// SIMATIC S7-200 project (STEP 7-Micro/WIN), CPU 224XP CN REL 02.01

SYMBOL_TABLE USUARIO1
C_1              VD100
C_0              VD110
L_k              VD180
r_k              VD190
m_k              VD120
m_k_1            VD130
m_k_2            VD140
e_k              VD300
e_k_1            VD160
e_k_2            VD170
Aa               VD200
Bb               VD210
Cc               VD220
Dd               VD230
Ee               VD240
r_k_1            VD250
END_SYMBOL_TABLE

ORGANIZATION_BLOCK PRINCIPAL:OB1
TITLE=COMENTARIOS DEL PROGRAMA
BEGIN
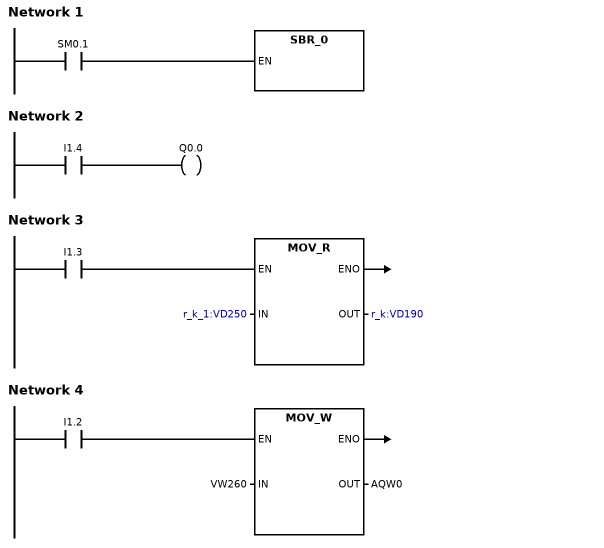
Network 1
LD     SM0.1
CALL   SBR_0:SBR0
Network 2
LD     I1.4
=      Q0.0
Network 3
LD     I1.3
MOVR   r_k_1:VD250, r_k:VD190
Network 4
LD     I1.2
MOVW   VW260, AQW0
END_ORGANIZATION_BLOCK

SUBROUTINE_BLOCK SBR_0:SBR0
TITLE=COMENTARIOS DE LA SUBRUTINA
BEGIN
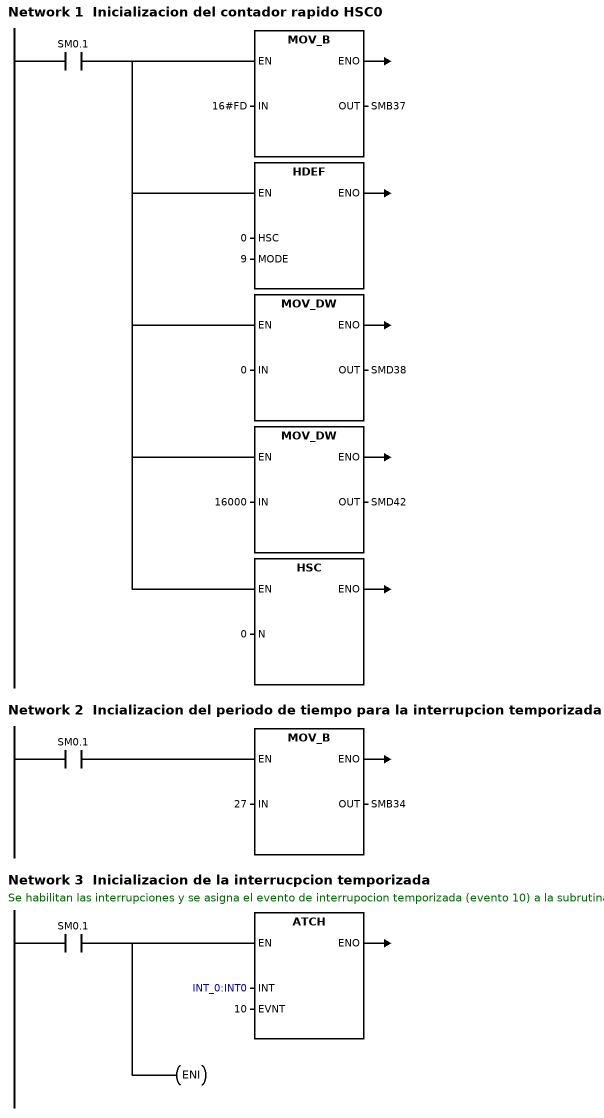
Network 1 // Inicializacion del contador rapido HSC0
LD     SM0.1
MOVB   16#FD, SMB37
HDEF   0, 9
MOVD   0, SMD38
MOVD   16000, SMD42
HSC    0
Network 2 // Incializacion del periodo de tiempo para la interrupcion temporizada
LD     SM0.1
MOVB   27, SMB34
Network 3 // Inicializacion de la interrucpcion temporizada
// Se habilitan las interrupciones y se asigna el evento de interrupocion temporizada (evento 10) a la subrutina de interrupcion INT_0
LD     SM0.1
ATCH   INT_0:INT0, 10
ENI
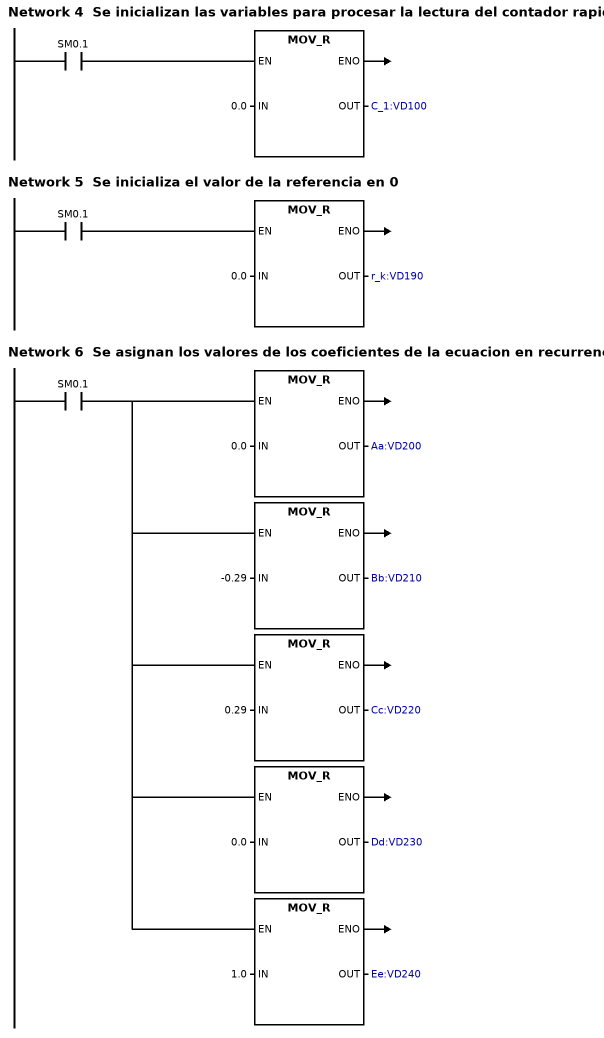
Network 4 // Se inicializan las variables para procesar la lectura del contador rapido HSC0
LD     SM0.1
MOVR   0.0, C_1:VD100
Network 5 // Se inicializa el valor de la referencia en 0
LD     SM0.1
MOVR   0.0, r_k:VD190
Network 6 // Se asignan los valores de los coeficientes de la ecuacion en recurrencia
LD     SM0.1
MOVR   0.0, Aa:VD200
MOVR   -0.29, Bb:VD210
MOVR   0.29, Cc:VD220
MOVR   0.0, Dd:VD230
MOVR   1.0, Ee:VD240
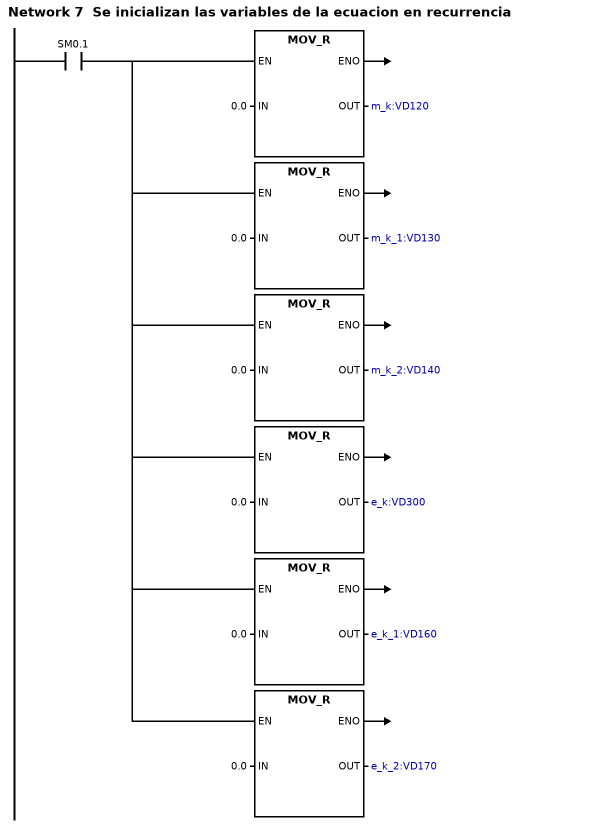
Network 7 // Se inicializan las variables de la ecuacion en recurrencia
LD     SM0.1
MOVR   0.0, m_k:VD120
MOVR   0.0, m_k_1:VD130
MOVR   0.0, m_k_2:VD140
MOVR   0.0, e_k:VD300
MOVR   0.0, e_k_1:VD160
MOVR   0.0, e_k_2:VD170
END_SUBROUTINE_BLOCK

INTERRUPT_BLOCK INT_0:INT0
TITLE=COMENTARIOS DE LA RUTINA DE INTERRUPCIÓN
BEGIN
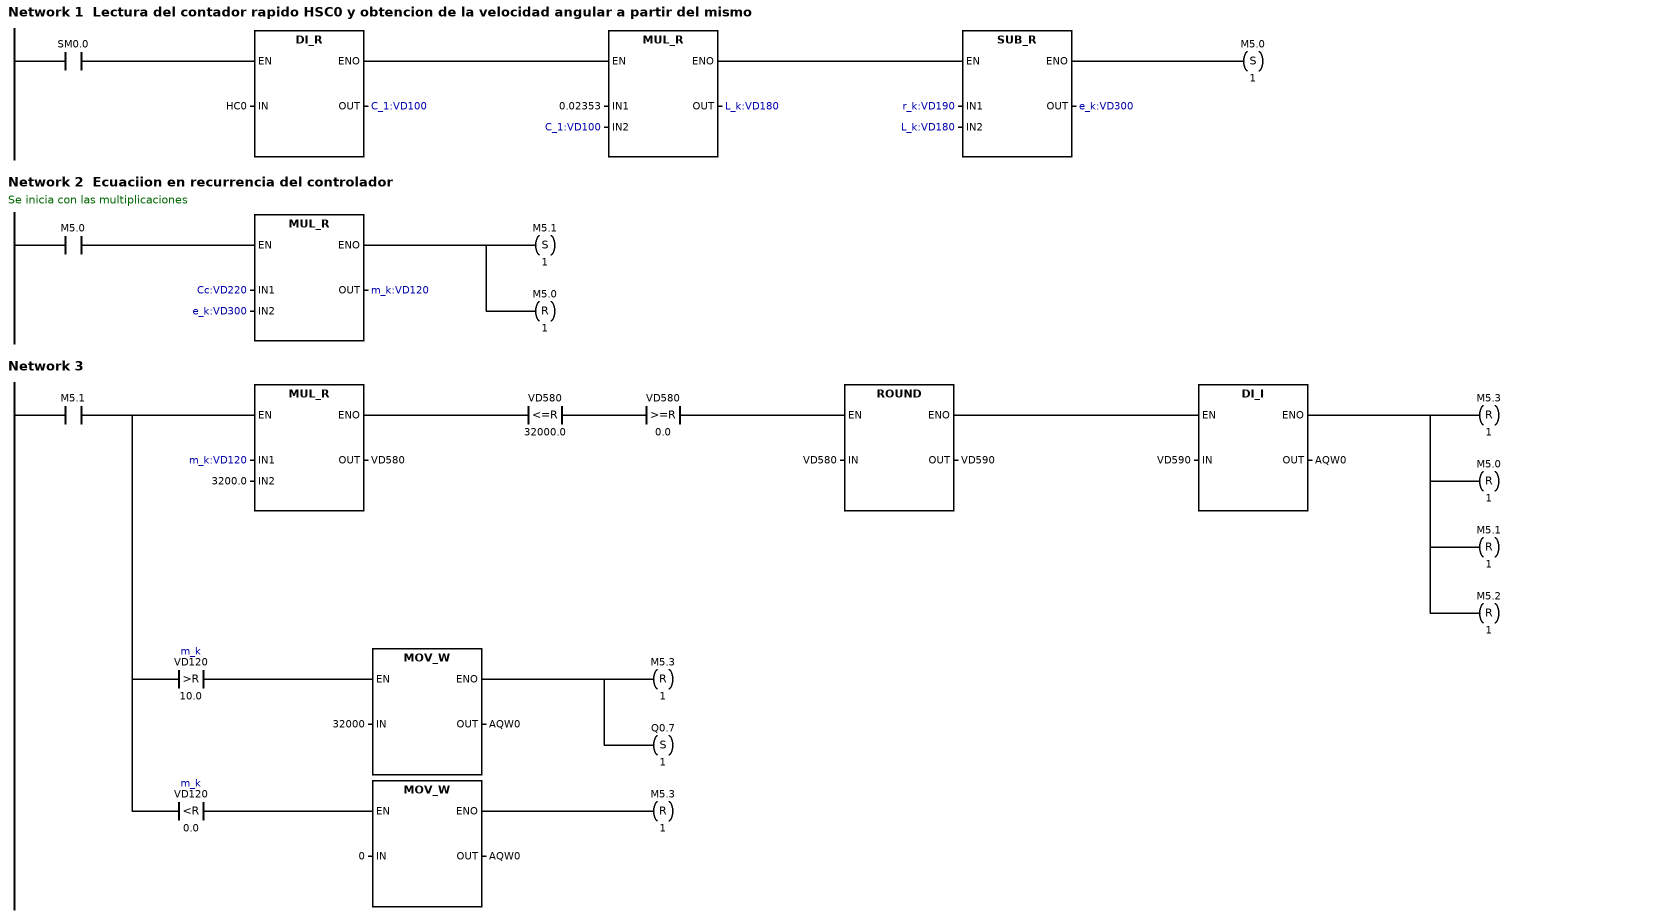
Network 1 // Lectura del contador rapido HSC0 y obtencion de la velocidad angular a partir del mismo
LD     SM0.0
DTR    HC0, C_1:VD100
AENO
MOVR   0.02353, L_k:VD180
AENO
*R     C_1:VD100, L_k:VD180
AENO
MOVR   r_k:VD190, e_k:VD300
AENO
-R     L_k:VD180, e_k:VD300
AENO
S      M5.0, 1
Network 2 // Ecuaciion en recurrencia del controlador 
// Se inicia con las multiplicaciones
LD     M5.0
MOVR   Cc:VD220, m_k:VD120
AENO
*R     e_k:VD300, m_k:VD120
AENO
S      M5.1, 1
R      M5.0, 1
Network 3
LD     M5.1
LPS
MOVR   m_k:VD120, VD580
AENO
*R     3200.0, VD580
AENO
AR<=   VD580, 32000.0
AR>=   VD580, 0.0
ROUND  VD580, VD590
AENO
DTI    VD590, AQW0
AENO
R      M5.3, 1
R      M5.0, 1
R      M5.1, 1
R      M5.2, 1
LRD
AR>    m_k:VD120, 10.0
MOVW   32000, AQW0
AENO
R      M5.3, 1
S      Q0.7, 1
LPP
AR<    m_k:VD120, 0.0
MOVW   0, AQW0
AENO
R      M5.3, 1
END_INTERRUPT_BLOCK
